// TIA Portal V20 export
// export: Created 2026-10-20T12:53:41.6428823Z, ExportSetting WithDefaults, DisplayName Totally Integrated Automation Portal, DisplayVersion V20 Update 6, DisplayName TIA Portal Openness, DisplayVersion V20 Update 6, DisplayName TIA Portal Version Control Interface, DisplayVersion V20 Update 6, DisplayName SINAMICS Startdrive Advanced, DisplayVersion V20 SP1, DisplayName SINAMICS Startdrive G130, G150, S120, S150, SINAMICS MV, G220, S200, S210, DisplayVersion V20 SP1, DisplayName SINAMICS Startdrive G110M, G120, G120C, G120D, G120P, G115D, DisplayVersion V20 SP1, DisplayName STEP 7 Professional, DisplayVersion V20 Update 6, DisplayName STEP 7 Safety, DisplayVersion V20 Update 2, DisplayName WinCC Basic/Comfort/Advanced, DisplayVersion V20 Update 6, DisplayName WinCC Unified, DisplayVersion V20 Update 6
DATA_BLOCK "Auto_Test_2_DB"   // DB118
VERSION : 0.1
// stored: AutoNumber true, DBAccessibleFromOPCUA true, InstanceOfName Auto_Test, InstanceOfType FB
"Auto_Test"
   // VAR_INPUT
   //    Sys_No : UInt;
   //    Automatic : Bool;
   //    Manual : Bool;
   //    Level : UInt;
   //    Error : Bool;
   //    Start : Bool;
   //    Pause : Bool;
   //    Stop : Bool;
   //    "Pallet Type" : Char;
   //    "Tower 1 Pallet Alignment" : Char;
   //    "Tower 2 Pallet Alignment" : Char;
   //    "Extractor Pallet Alignment" : Char;
   //    Pallet_Allignment : Char;
   //    Tower : UInt;
   //    Transfer_From_To : Byte;
   //    "From level" : Byte;
   //    "To level" : Byte;
   //    "Testing Time" : UInt;
   //    "Numer of cycles" : Byte;
   // END_VAR
   // VAR_OUTPUT
   //    Running : Bool;
   //    Time_Runnng : Time;
   //    Start_Time { ExternalAccessible := 'False'; ExternalVisible := 'False'; ExternalWritable := 'False'} : String;
   //    Stop_Time { ExternalAccessible := 'False'; ExternalVisible := 'False'; ExternalWritable := 'False'} : String;
   //    Duration : Time;
   // END_VAR
   // VAR_IN_OUT
   //    "Order Table_1" : "OrderTable_UDT";
   //    Step_Table_0 : "OrderTable_UDT";
   //    System_OrderSent : Bool;
   //    Total_Duration : Time;
   // END_VAR
   // VAR
   //    State : Int;
   //    R_Start { S7_SetPoint := 'True'} : R_TRIG;
   //    T_Delay { S7_SetPoint := 'True'} : TON_TIME;
   //    Time_Delay : Time;
   //    Send_VTD_Order : Bool;
   //    Send_CNV_Order : Bool;
   //    R_TRIG_Instance { S7_SetPoint := 'True'} : R_TRIG;
   //    T_Running { S7_SetPoint := 'True'} : TON_TIME;
   //    F_TRIG { S7_SetPoint := 'True'} : F_TRIG;
   //    R_TRIG { S7_SetPoint := 'True'} : R_TRIG;
   //    Error_Code : Int;
   //    test : Bool;
   //    N_Cycles : UInt;
   //    Testing_Time : Time;
   //    R_Manual_Mode { S7_SetPoint := 'True'} : R_TRIG;
   // END_VAR
BEGIN
END_DATA_BLOCK
